Fanuc KAREL source: kd00024.KL

-- PROVISIONAL review KL for V1013-1; original PC SHA256 6ee5e4d0683bfa0b2830b7f5e70fafd68b5e58b162bae63cc5a37ee6ab8760a1
-- Incomplete behavior may be omitted. Consult companion uncertainty JSON. Do not deploy.
PROGRAM KD00024
%NOLOCKGROUP
VAR
  I : INTEGER
  J : INTEGER
  B : BOOLEAN
  R : REAL
  S : STRING[80]
BEGIN
  -- UNRESOLVED_PC offsets 5-12; opcodes 9D,23
  -- UNRESOLVED_PC offsets 17-50; opcodes 9D,81,18,22,2E,21,54,12,22,9D,13,04
  -- UNRESOLVED_PC offsets 55-59; opcodes 7F
END KD00024
